(* CODESYS project ASRS_RLI_Presse.project

Project tree, tasks and I/O mapping:
  PLCWinNT : CODESYS Control Win V3, CODESYS, version 3.5.22.40
    application Application
      libraries: Standard, * (System)
      task MainTask (cyclic, interval 10 ms, priority 1) calls PLC_PRG
      task VISU_TASK (cyclic, interval 100 ms, priority 31) calls VisuElems.Visu_Prg
      program PLC_PRG [ST]
      function block FB_RLI_Presse [ST]
      function block FB_RLI_PresseTests [ST]
      visualisation VISU_RLI_PRESSE
  text list GlobalTextList
*)

// PLCWinNT/Application/PLC_PRG
PROGRAM PLC_PRG
VAR
    Press : FB_RLI_Presse;
    StartRequest : BOOL;
    ReleaseRequest : BOOL;
    ResetFault : BOOL;
    StationEnabled : BOOL := TRUE;
    HoldPress : BOOL;
    ReplayReply : BOOL;
    Tests : FB_RLI_PresseTests;
    StateText : STRING(48);
    FaultText : STRING(55);
END_VAR

Press(
    StartRequest := StartRequest,
    ReleaseRequest := ReleaseRequest,
    ResetFault := ResetFault,
    StationEnabled := StationEnabled,
    HoldPress := HoldPress,
    ReplayReply := ReplayReply
);
StartRequest := FALSE;
ReleaseRequest := FALSE;
ResetFault := FALSE;
Tests();

CASE Press.State OF
    0: StateText := 'En attente';
    10: StateText := 'Confirmation presse attendue';
    20: StateText := 'Autorisation de transfert simulee';
    90: StateText := 'Defaut verrouille';
ELSE
    StateText := 'Etat inconnu';
END_CASE;

CASE Press.FaultCode OF
    0: FaultText := 'Aucun';
    1: FaultText := 'Echanges station perimes';
    2: FaultText := 'Delai de commande depasse';
ELSE
    FaultText := 'Code non identifie';
END_CASE;

END_PROGRAM

// PLCWinNT/Application/FB_RLI_Presse
FUNCTION_BLOCK FB_RLI_Presse
VAR_INPUT
    StartRequest : BOOL;
    ReleaseRequest : BOOL;
    ResetFault : BOOL;
    StationEnabled : BOOL := TRUE;
    HoldPress : BOOL;
    ReplayReply : BOOL;
END_VAR
VAR_OUTPUT
    State : USINT;
    FaultCode : USINT;
    LinkFresh : BOOL;
    TransferAllowed : BOOL;
    StaleReply : BOOL;
    ReplyValid : BOOL;
    RequestId : UINT;
    ReplyId : UINT;
    Tx : ARRAY[0..3] OF BYTE;
    Rx : ARRAY[0..3] OF BYTE;
END_VAR
VAR
    StartEdge : R_TRIG;
    ReleaseEdge : R_TRIG;
    ResetEdge : R_TRIG;
    HeartbeatPeriod : TON;
    Watchdog : TON;
    PressDelay : TON;
    CommandDeadline : TON;
    Heartbeat : BYTE;
    PreviousHeartbeat : BYTE;
    HeartbeatChanges : USINT;
    HeartbeatChanged : BOOL;
    LinkWasReady : BOOL;
    TxRequestId : UINT;
    LastReplyId : UINT;
    LastReplyValid : BOOL;

    ReplyStopped : BOOL;
END_VAR

// A virtual station consumes the output image from the preceding scan.
// Its input image freezes when the station is disabled.
HeartbeatPeriod(IN := StationEnabled AND NOT HeartbeatPeriod.Q, PT := T#100ms);
PressDelay(IN := StationEnabled AND (Tx[0] = BYTE#1) AND NOT HoldPress AND NOT ReplayReply,
           PT := T#400ms);
IF StationEnabled THEN
    IF HeartbeatPeriod.Q THEN
        IF Heartbeat = BYTE#255 THEN
            Heartbeat := BYTE#0;
        ELSE
            Heartbeat := Heartbeat + BYTE#1;
        END_IF;
    END_IF;
    Rx[1] := Heartbeat;
    TxRequestId := BYTE_TO_UINT(Tx[2]) + BYTE_TO_UINT(Tx[3]) * UINT#256;
    Rx[0] := BYTE#0;
    IF ReplayReply AND LastReplyValid THEN
        Rx[0] := BYTE#3;
        Rx[2] := UINT_TO_BYTE(LastReplyId MOD UINT#256);
        Rx[3] := UINT_TO_BYTE(LastReplyId / UINT#256);
    ELSIF PressDelay.Q THEN
        LastReplyId := TxRequestId;
        LastReplyValid := TRUE;
        Rx[0] := BYTE#3;
        Rx[2] := Tx[2];
        Rx[3] := Tx[3];
    END_IF;
END_IF;

// The watchdog consumes the image only. StationEnabled is a bench stimulus.
HeartbeatChanged := Rx[1] <> PreviousHeartbeat;
PreviousHeartbeat := Rx[1];
Watchdog(IN := NOT HeartbeatChanged, PT := T#350ms);
IF Watchdog.Q THEN
    HeartbeatChanges := USINT#0;
ELSIF HeartbeatChanged AND (HeartbeatChanges < USINT#2) THEN
    HeartbeatChanges := HeartbeatChanges + USINT#1;
END_IF;
LinkFresh := HeartbeatChanges = USINT#2;
IF LinkFresh THEN
    LinkWasReady := TRUE;
END_IF;

ReplyValid := (Rx[0] AND BYTE#1) <> BYTE#0;
ReplyStopped := (Rx[0] AND BYTE#2) <> BYTE#0;
ReplyId := BYTE_TO_UINT(Rx[2]) + BYTE_TO_UINT(Rx[3]) * UINT#256;
StaleReply := LinkFresh AND (State = USINT#10 OR State = USINT#20)
              AND ReplyValid AND (ReplyId <> RequestId);

StartEdge(CLK := StartRequest);
ReleaseEdge(CLK := ReleaseRequest);
ResetEdge(CLK := ResetFault);
CommandDeadline(IN := State = USINT#10, PT := T#2s);

IF LinkWasReady AND NOT LinkFresh AND State <> USINT#90 THEN
    FaultCode := USINT#1;
    State := USINT#90;
ELSE
    CASE State OF
        0:
            IF LinkFresh AND StartEdge.Q THEN
                IF RequestId = UINT#65535 THEN
                    RequestId := UINT#1;
                ELSE
                    RequestId := RequestId + UINT#1;
                END_IF;
                State := USINT#10;
            END_IF;
        10:
            IF CommandDeadline.Q THEN
                FaultCode := USINT#2;
                State := USINT#90;
            ELSIF LinkFresh AND ReplyValid AND ReplyStopped AND (ReplyId = RequestId) THEN
                State := USINT#20;
            END_IF;
        20:
            IF NOT ReplyValid OR NOT ReplyStopped OR (ReplyId <> RequestId) THEN
                FaultCode := USINT#3;
                State := USINT#90;
            ELSIF ReleaseEdge.Q THEN
                State := USINT#0;
            END_IF;
        90:
            IF LinkFresh AND ResetEdge.Q AND NOT StartRequest THEN
                FaultCode := USINT#0;
                State := USINT#0;
            END_IF;
    END_CASE;
END_IF;

TransferAllowed := (State = USINT#20) AND LinkFresh;
IF State = USINT#10 OR State = USINT#20 THEN
    Tx[0] := BYTE#1;
ELSE
    Tx[0] := BYTE#0;
END_IF;
Tx[1] := BYTE#0; // Reserved.
Tx[2] := UINT_TO_BYTE(RequestId MOD UINT#256);
Tx[3] := UINT_TO_BYTE(RequestId / UINT#256);

END_FUNCTION_BLOCK

// PLCWinNT/Application/FB_RLI_PresseTests
FUNCTION_BLOCK FB_RLI_PresseTests
VAR_OUTPUT
    Done : BOOL;
    Passed : BOOL;
    FailedCase : USINT;
    TestStage : USINT;
END_VAR
VAR
    Bench : FB_RLI_Presse;
    StageAge : TON;
    PreviousStage : USINT := USINT#255;
    OldRequest : UINT;
END_VAR

// Use a separate bench instance so acceptance tests do not change operator inputs.
StageAge(IN := TestStage = PreviousStage, PT := T#4s);
PreviousStage := TestStage;

Bench(
    StartRequest := (TestStage = USINT#10) OR (TestStage = USINT#30)
                    OR (TestStage = USINT#50) OR (TestStage = USINT#70)
                    OR (TestStage = USINT#80) OR (TestStage = USINT#81) OR (TestStage = USINT#84),
    ReleaseRequest := TestStage = USINT#20,
    ResetFault := (TestStage = USINT#40) OR (TestStage = USINT#60)
                  OR (TestStage = USINT#81) OR (TestStage = USINT#83),
    StationEnabled := TestStage <> USINT#80,
    HoldPress := TestStage = USINT#50,
    ReplayReply := TestStage = USINT#30
);

IF NOT Done THEN
    CASE TestStage OF
        0: // Wait until the station has sent two distinct heartbeats.
            IF Bench.LinkFresh THEN
                TestStage := USINT#10;
            END_IF;
        10: // Nominal stop request, correlated confirmation and permit.
            IF Bench.TransferAllowed AND (Bench.ReplyId = Bench.RequestId)
               AND (Bench.RequestId <> UINT#0) THEN
                OldRequest := Bench.RequestId;
                TestStage := USINT#20;
            END_IF;
        20:
            IF (Bench.State = USINT#0) AND NOT Bench.TransferAllowed THEN
                TestStage := USINT#30;
            END_IF;
        30: // Replay the previous completed request while the station stays live.
            IF Bench.TransferAllowed OR NOT Bench.LinkFresh THEN
                FailedCase := TestStage;
            ELSIF Bench.FaultCode = USINT#2 THEN
                IF Bench.ReplyId = OldRequest AND Bench.RequestId <> OldRequest THEN
                    TestStage := USINT#40;
                ELSE
                    FailedCase := TestStage;
                END_IF;
            END_IF;
        40:
            IF Bench.State = USINT#0 THEN
                TestStage := USINT#50;
            END_IF;
        50: // Live station with no completion response.
            IF Bench.TransferAllowed OR NOT Bench.LinkFresh THEN
                FailedCase := TestStage;
            ELSIF Bench.FaultCode = USINT#2 THEN
                TestStage := USINT#60;
            END_IF;
        60:
            IF Bench.State = USINT#0 THEN
                TestStage := USINT#70;
            END_IF;
        70: // Obtain a permit again before interrupting the link.
            IF Bench.TransferAllowed THEN
                TestStage := USINT#80;
            END_IF;
        80: // Freeze last image, then require the watchdog to revoke the permit.
            IF Bench.FaultCode = USINT#1 THEN
                IF NOT Bench.TransferAllowed AND NOT Bench.LinkFresh THEN
                    TestStage := USINT#81;
                ELSE
                    FailedCase := TestStage;
                END_IF;
            END_IF;
        81: // Reconnect while both start and reset are already held.
            IF Bench.TransferAllowed OR (Bench.State <> USINT#90) THEN
                FailedCase := TestStage;
            ELSIF Bench.LinkFresh THEN
                TestStage := USINT#82;
            END_IF;
        82: // Release both before requesting an explicit reset.
            IF (Bench.State = USINT#90) AND NOT Bench.TransferAllowed THEN
                TestStage := USINT#83;
            ELSE
                FailedCase := TestStage;
            END_IF;
        83: // Reset returns to idle without granting the transfer.
            IF Bench.State = USINT#0 AND NOT Bench.TransferAllowed THEN
                OldRequest := Bench.RequestId;
                TestStage := USINT#84;
            END_IF;
        84: // A fresh start is required and must allocate a new request ID.
            IF Bench.TransferAllowed AND (Bench.RequestId <> OldRequest) THEN
                TestStage := USINT#100;
                Passed := TRUE;
                Done := TRUE;
            END_IF;
    END_CASE;
    IF StageAge.Q OR FailedCase <> USINT#0 THEN
        // Stage 0 has no case number, so code 1 denotes initial-link failure.
        IF FailedCase = USINT#0 THEN
            IF TestStage = USINT#0 THEN
                FailedCase := USINT#1;
            ELSE
                FailedCase := TestStage;
            END_IF;
        END_IF;
        Done := TRUE;
        Passed := FALSE;
    END_IF;
END_IF;

END_FUNCTION_BLOCK

// PLCWinNT/Application/VISU_RLI_PRESSE
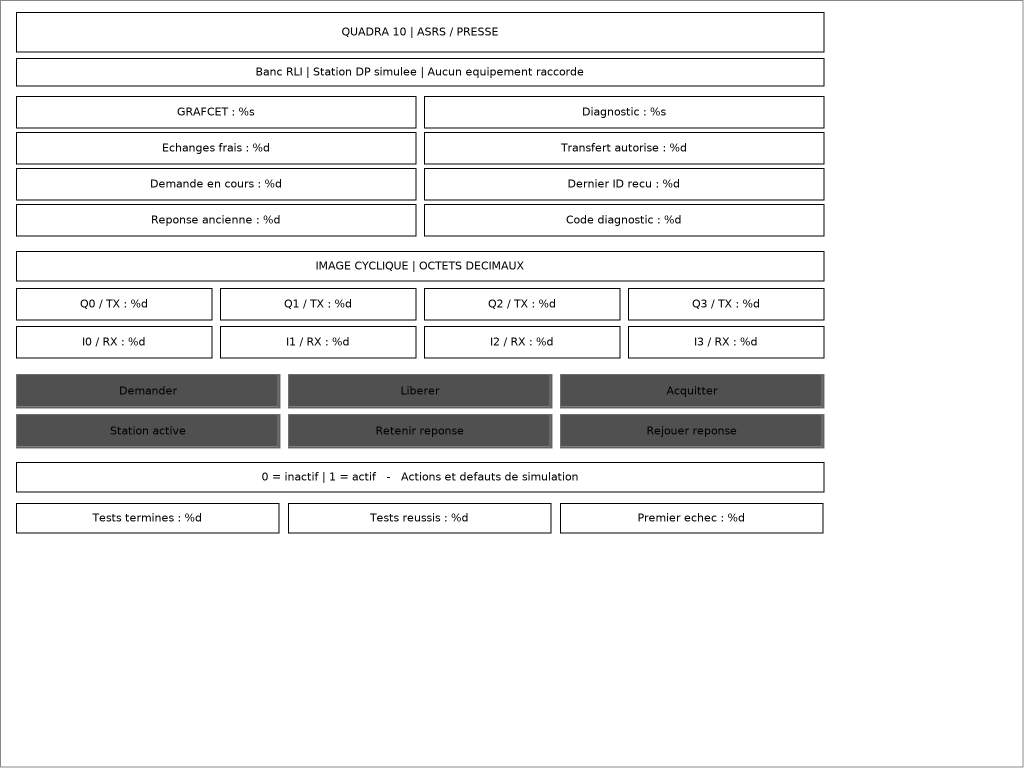
VISUALIZATION VISU_RLI_PRESSE  // 1024x768
    Rectangle (16,12 808x40), "QUADRA 10 | ASRS / PRESSE"
    Rectangle (16,58 808x28), "Banc RLI | Station DP simulee | Aucun equipement raccorde"
    Rectangle (16,96 400x32), "GRAFCET : %s", text variable: PLC_PRG.StateText
    Rectangle (424,96 400x32), "Diagnostic : %s", text variable: PLC_PRG.FaultText
    Rectangle (16,132 400x32), "Echanges frais : %d", text variable: PLC_PRG.Press.LinkFresh
    Rectangle (424,132 400x32), "Transfert autorise : %d", text variable: PLC_PRG.Press.TransferAllowed
    Rectangle (16,168 400x32), "Demande en cours : %d", text variable: PLC_PRG.Press.RequestId
    Rectangle (424,168 400x32), "Dernier ID recu : %d", text variable: PLC_PRG.Press.ReplyId
    Rectangle (16,204 400x32), "Reponse ancienne : %d", text variable: PLC_PRG.Press.StaleReply
    Rectangle (424,204 400x32), "Code diagnostic : %d", text variable: PLC_PRG.Press.FaultCode
    Rectangle (16,251 808x30), "IMAGE CYCLIQUE | OCTETS DECIMAUX"
    Rectangle (16,288 196x32), "Q0 / TX : %d", text variable: PLC_PRG.Press.Tx[0]
    Rectangle (16,326 196x32), "I0 / RX : %d", text variable: PLC_PRG.Press.Rx[0]
    Rectangle (220,288 196x32), "Q1 / TX : %d", text variable: PLC_PRG.Press.Tx[1]
    Rectangle (220,326 196x32), "I1 / RX : %d", text variable: PLC_PRG.Press.Rx[1]
    Rectangle (424,288 196x32), "Q2 / TX : %d", text variable: PLC_PRG.Press.Tx[2]
    Rectangle (424,326 196x32), "I2 / RX : %d", text variable: PLC_PRG.Press.Rx[2]
    Rectangle (628,288 196x32), "Q3 / TX : %d", text variable: PLC_PRG.Press.Tx[3]
    Rectangle (628,326 196x32), "I3 / RX : %d", text variable: PLC_PRG.Press.Rx[3]
    Button (16,374 264x34), "Demander"
        OnMouseClick: execute { PLC_PRG.StartRequest := TRUE; }
    Button (288,374 264x34), "Liberer"
        OnMouseClick: execute { PLC_PRG.ReleaseRequest := TRUE; }
    Button (560,374 264x34), "Acquitter"
        OnMouseClick: execute { PLC_PRG.ResetFault := TRUE; }
    Button (16,414 264x34), "Station active"
        OnMouseClick: execute { PLC_PRG.StationEnabled := NOT PLC_PRG.StationEnabled; }
    Button (288,414 264x34), "Retenir reponse"
        OnMouseClick: execute { PLC_PRG.HoldPress := NOT PLC_PRG.HoldPress; }
    Button (560,414 264x34), "Rejouer reponse"
        OnMouseClick: execute { PLC_PRG.ReplayReply := NOT PLC_PRG.ReplayReply; }
    Rectangle (16,462 808x30), "0 = inactif | 1 = actif - Actions et defauts de simulation"
    Rectangle (16,503 263x30), "Tests termines : %d", text variable: PLC_PRG.Tests.Done
    Rectangle (288,503 263x30), "Tests reussis : %d", text variable: PLC_PRG.Tests.Passed
    Rectangle (560,503 263x30), "Premier echec : %d", text variable: PLC_PRG.Tests.FailedCase
END_VISUALIZATION
